(* PLC project minimal, x x 1 *)
(* stored: creationDateTime 2026-01-01T00:00:00 *)

PROGRAM drive
  VAR_OUTPUT
    A : BOOL;
    B : BOOL;
  END_VAR

A := TRUE;
B := TRUE;
END_PROGRAM

CONFIGURATION C
  RESOURCE R ON PLC
    TASK t(INTERVAL := T#10ms, PRIORITY := 0);
    PROGRAM i WITH t : drive;
  END_RESOURCE
END_CONFIGURATION
